(* IEC 61131-3 sources: ZPLC/packages/zplc-ide/projects/il_interlock_guard/src, 1 file *)

(* ---- MotorPlant.il ---- *)
PROGRAM MotorPlant
VAR_INPUT
    Start AT %I0.0 : BOOL;
    Stop AT %I0.1 : BOOL;
    AtSpeed AT %I0.2 : BOOL;
    GuardClosed AT %I0.3 : BOOL;
END_VAR
VAR_OUTPUT
    Command AT %Q0.0 : BOOL;
    Running AT %Q0.1 : BOOL;
END_VAR

        LD    Start
        OR    Command
        ANDN  Stop
        AND   GuardClosed
        ST    Command
        AND   AtSpeed
        ST    Running
END_PROGRAM
